(* Logix 5000 project; controller TFF vendor 1 type 14 code 107 rev 33.11; software revision 33.04; part 33 of 38 *)
(* tags used below, declared in another part *)
   Address : DINT;   // Temp Address
   Index : DINT;   // Index
   Index2 : DINT;   // Index
   result : DINT[2];
   SCL : SCALE;   // Scale Instruction
   AlarmAnalog : AlarmAnalog[50];   // Analog Alarm Array
   AlarmControl : AlarmControl;   // Alarm Control
   AnalogOutput : AnalogOutput[25];   // Analog Output Array
   AnalogPoint : AnalogInput[50];   // Analog Input Array
   DigitalInput : BOOL[256];   // Digital Input Array these bits are copied from Input cards.
   DigitalPoint : DigitalPoint[150];   // Digital Point Array
   ES001 : ALIAS FOR DigitalPoint[2];
   FlowPath : FlowPath[64];   // Flow Path Array
   FlowPathControl : FlowPathControl;   // Flow Path Control
   RawAnalogInputArray : INT[50];   // Array of analog input raw
   SysControl : SysControl;   // General system status and command
   Valve : Valve[100];   // Valve Array
   ValveControl : ValveControl;   // Valve Control
   ValveSwInput : BOOL[64];   // Valve digital input
(* Process, continued *)

ROUTINE modInputAnalog   (* ladder *)
// Analog Input Routine
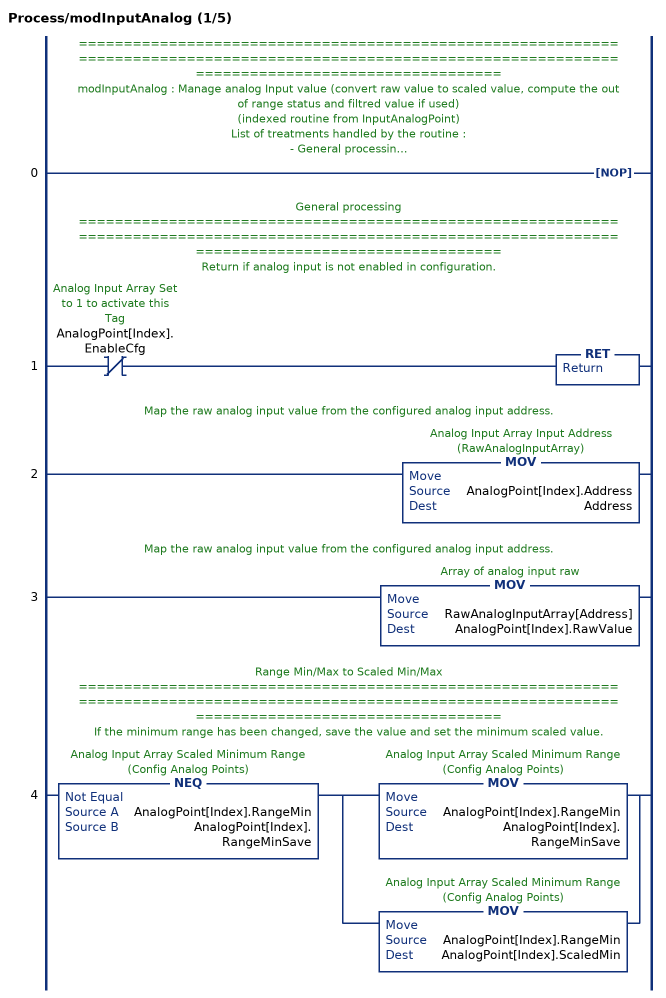
   // ==========================================================================================================================================================
   //                                            modInputAnalog : Manage analog Input value (convert raw value to scaled value, compute the out of range status and filtred value if used)
   //                                                                                                                        (indexed routine from InputAnalogPoint)
   //                                                     List of treatments handled by the routine :
   //                                                          - General processing
   //                                                          - Range Min/Max to Scaled Min/Max
   //                                                          - Out of Range status calculation
   //                                                          - filtering raw value
   //                                                          - Compute scaled value
   //                                                          - Map analog input value to alarm analog value
   //                                                     -----------------------------------------------------------------------------------------------------------------------------------------------------
   //                                                     History
   // 		2019-DEC-24 - Merck - Q. Spindler - Initial version for Candidate Release 1.00.00.00.a
   // 		2021-MAY-21 - Merck - Q. Spindler - Modifications for Candidate Release 1.00.00.00.e
   //                                                     - Out of Range status calculation, add exception for pressure sensors
   // ==========================================================================================================================================================
   0: NOP();
   // General processing
   // ==========================================================================================================================================================
   // Return if analog input is not enabled in configuration.
   1: XIO(AnalogPoint[Index].EnableCfg)RET();
   // Map the raw analog input value from the configured analog input address.
   2: MOV(AnalogPoint[Index].Address,Address);
   // Map the raw analog input value from the configured analog input address.
   3: MOV(RawAnalogInputArray[Address],AnalogPoint[Index].RawValue);
   // Range Min/Max to Scaled Min/Max
   // ==========================================================================================================================================================
   // If the minimum range has been changed, save the value and set the minimum scaled value.
   4: NEQ(AnalogPoint[Index].RangeMin,AnalogPoint[Index].RangeMinSave)[MOV(AnalogPoint[Index].RangeMin,AnalogPoint[Index].RangeMinSave) ,MOV(AnalogPoint[Index].RangeMin,AnalogPoint[Index].ScaledMin) ];
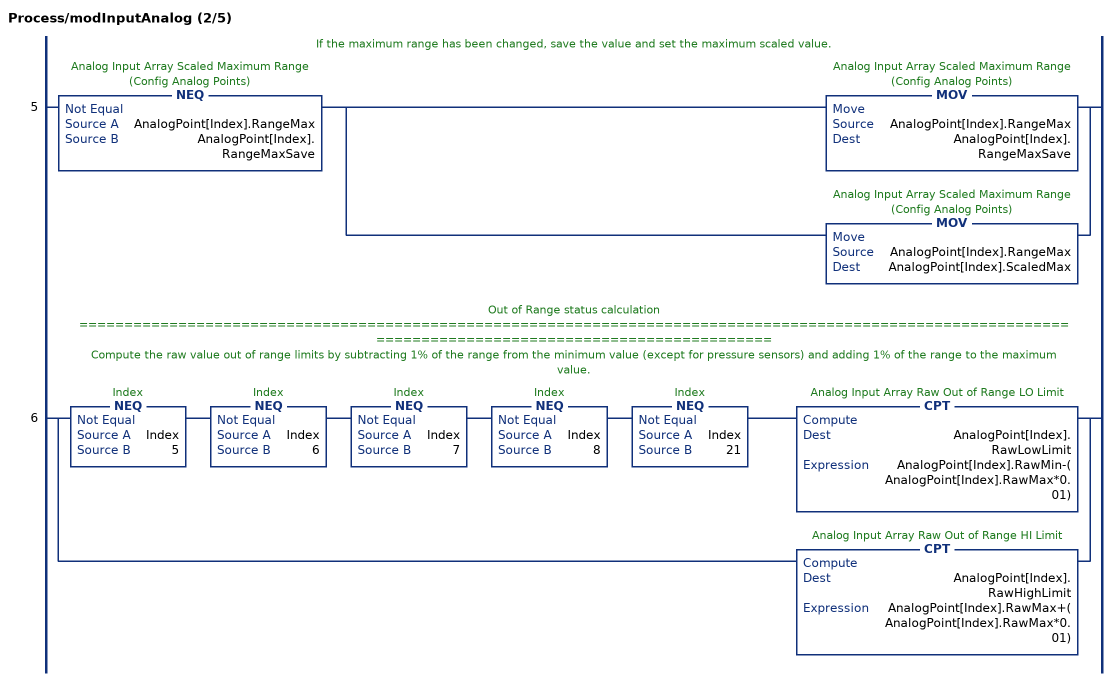
   // If the maximum range has been changed, save the value and set the maximum scaled value.
   5: NEQ(AnalogPoint[Index].RangeMax,AnalogPoint[Index].RangeMaxSave)[MOV(AnalogPoint[Index].RangeMax,AnalogPoint[Index].RangeMaxSave) ,MOV(AnalogPoint[Index].RangeMax,AnalogPoint[Index].ScaledMax) ];
   // Out of Range status calculation
   // ==========================================================================================================================================================
   // Compute the raw value out of range limits by subtracting 1% of the range from the minimum value (except for pressure sensors) and adding 1% of the range to the maximum value.
   6: [NEQ(Index,5) NEQ(Index,6) NEQ(Index,7) NEQ(Index,8) NEQ(Index,21) CPT(AnalogPoint[Index].RawLowLimit,AnalogPoint[Index].RawMin-(AnalogPoint[Index].RawMax*0.01)) ,CPT(AnalogPoint[Index].RawHighLimit,AnalogPoint[Index].RawMax+(AnalogPoint[Index].RawMax*0.01)) ];
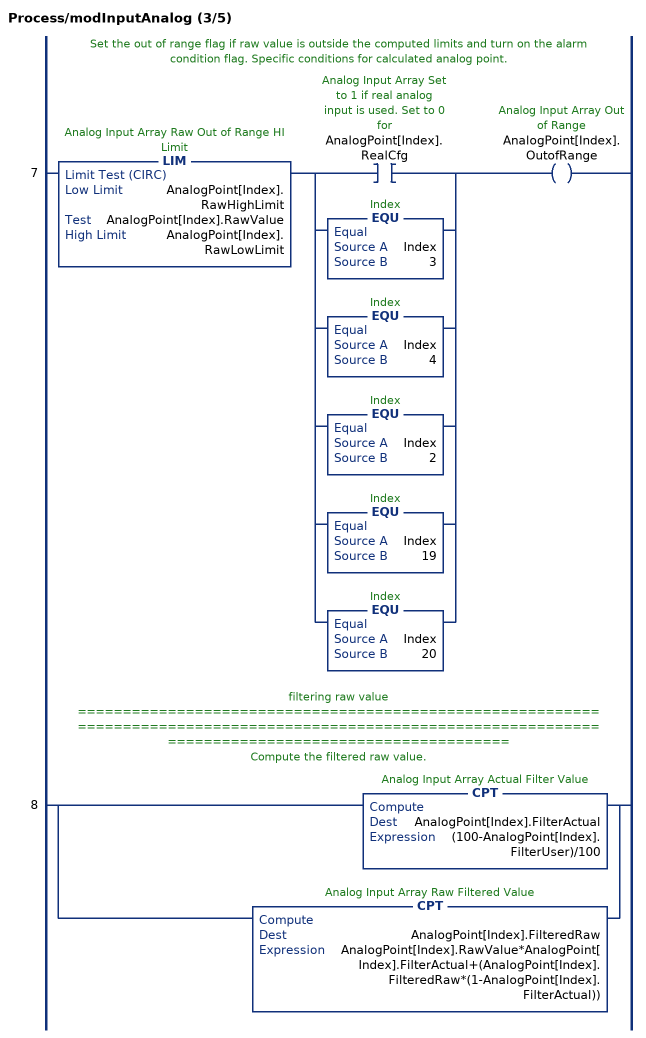
   // Set the out of range flag if raw value is outside the computed limits and turn on the alarm condition flag. Specific conditions for calculated analog point.
   7: LIM(AnalogPoint[Index].RawHighLimit,AnalogPoint[Index].RawValue,AnalogPoint[Index].RawLowLimit)[XIC(AnalogPoint[Index].RealCfg) ,EQU(Index,3) ,EQU(Index,4) ,EQU(Index,2) ,EQU(Index,19) ,EQU(Index,20) ]OTE(AnalogPoint[Index].OutofRange);
   // filtering raw value
   // ==========================================================================================================================================================
   // Compute the filtered raw value.
   8: [CPT(AnalogPoint[Index].FilterActual,(100-AnalogPoint[Index].FilterUser)/100) ,CPT(AnalogPoint[Index].FilteredRaw,AnalogPoint[Index].RawValue*AnalogPoint[Index].FilterActual+(AnalogPoint[Index].FilteredRaw*(1-AnalogPoint[Index].FilterActual))) ];
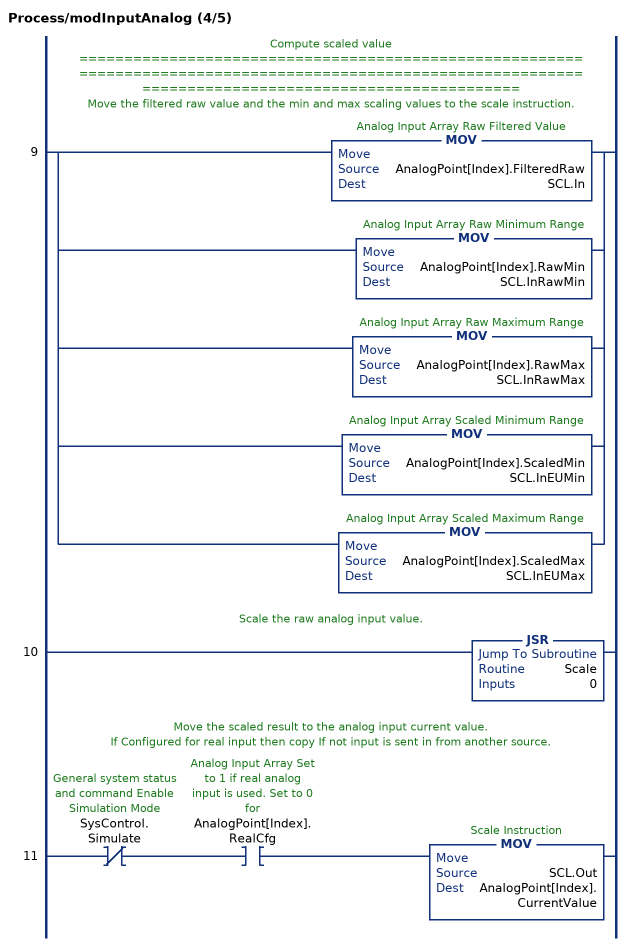
   // Compute scaled value
   // ==========================================================================================================================================================
   // Move the filtered raw value and the min and max scaling values to the scale instruction.
   9: [MOV(AnalogPoint[Index].FilteredRaw,SCL.In) ,MOV(AnalogPoint[Index].RawMin,SCL.InRawMin) ,MOV(AnalogPoint[Index].RawMax,SCL.InRawMax) ,MOV(AnalogPoint[Index].ScaledMin,SCL.InEUMin) ,MOV(AnalogPoint[Index].ScaledMax,SCL.InEUMax) ];
   // Scale the raw analog input value.
   10: JSR(Scale,0);
   // Move the scaled result to the analog input current value.
   // If Configured for real input then copy If not input is sent in from another source.
   11: XIO(SysControl.Simulate)XIC(AnalogPoint[Index].RealCfg)MOV(SCL.Out,AnalogPoint[Index].CurrentValue);
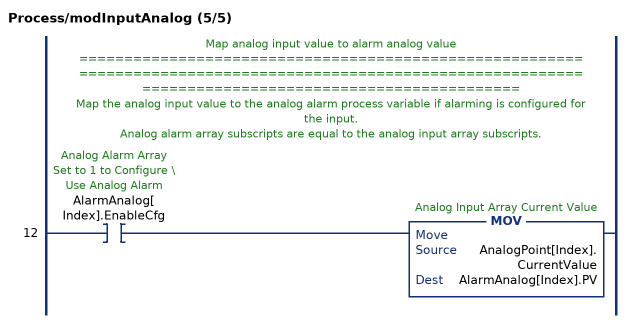
   // Map analog input value to alarm analog value
   // ==========================================================================================================================================================
   // Map the analog input value to the analog alarm process variable if alarming is configured for the input.
   // Analog alarm array subscripts are equal to the analog input array subscripts.
   12: XIC(AlarmAnalog[Index].EnableCfg)MOV(AnalogPoint[Index].CurrentValue,AlarmAnalog[Index].PV);
END_ROUTINE

ROUTINE modInputDigital   (* ladder *)
// Digital Input Routine
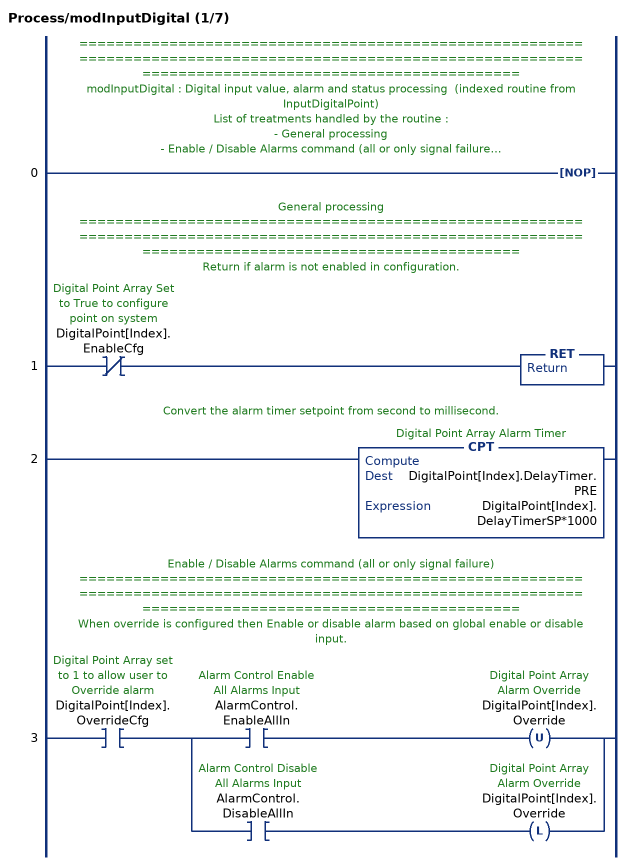
   // ==========================================================================================================================================================
   //                                                        modInputDigital : Digital input value, alarm and status processing  (indexed routine from InputDigitalPoint)
   //                                                     List of treatments handled by the routine :
   //                                                          - General processing
   //                                                          - Enable / Disable Alarms command (all or only signal failure)
   //                                                          - Digital alarm processing
   //                                                          - Digital input status
   //                                                          - Digital alarm status acknowledged
   //                                                          - Digital alarm status
   //                                                          - General processing
   //                                                          - Compute current value
   //                                                     -----------------------------------------------------------------------------------------------------------------------------------------------------
   //                                                     History
   // 		2019-DEC-24 - Merck - Q. Spindler - Initial version for Candidate Release 1.00.00.00.a
   // ==========================================================================================================================================================
   0: NOP();
   // General processing
   // ==========================================================================================================================================================
   // Return if alarm is not enabled in configuration.
   1: XIO(DigitalPoint[Index].EnableCfg)RET();
   // Convert the alarm timer setpoint from second to millisecond.
   2: CPT(DigitalPoint[Index].DelayTimer.PRE,DigitalPoint[Index].DelayTimerSP*1000);
   // Enable / Disable Alarms command (all or only signal failure)
   // ==========================================================================================================================================================
   // When override is configured then Enable or disable alarm based on global enable or disable input.
   3: XIC(DigitalPoint[Index].OverrideCfg)[XIC(AlarmControl.EnableAllIn) OTU(DigitalPoint[Index].Override) ,XIC(AlarmControl.DisableAllIn) OTL(DigitalPoint[Index].Override) ];
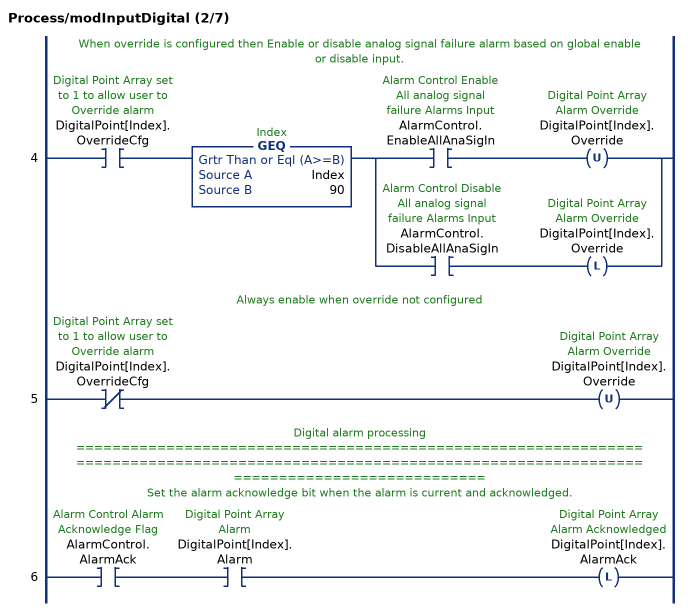
   // When override is configured then Enable or disable analog signal failure alarm based on global enable or disable input.
   4: XIC(DigitalPoint[Index].OverrideCfg)GEQ(Index,90)[XIC(AlarmControl.EnableAllAnaSigIn) OTU(DigitalPoint[Index].Override) ,XIC(AlarmControl.DisableAllAnaSigIn) OTL(DigitalPoint[Index].Override) ];
   // Always enable when override not configured
   5: XIO(DigitalPoint[Index].OverrideCfg)OTU(DigitalPoint[Index].Override);
   // Digital alarm processing
   // ==========================================================================================================================================================
   // Set the alarm acknowledge bit when the alarm is current and acknowledged.
   6: XIC(AlarmControl.AlarmAck)XIC(DigitalPoint[Index].Alarm)OTL(DigitalPoint[Index].AlarmAck);
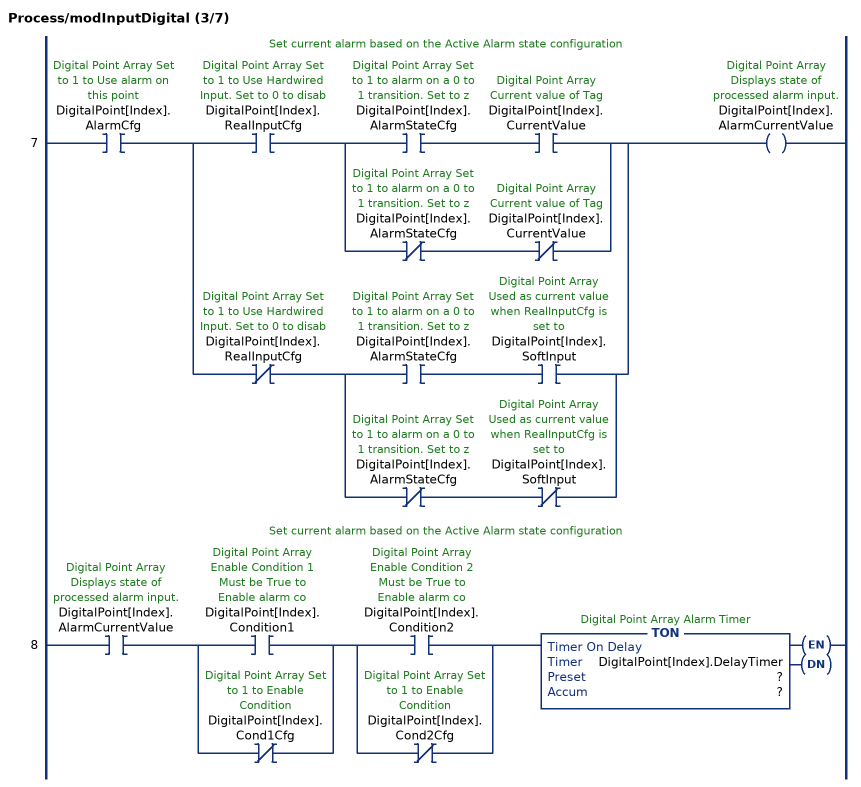
   // Set current alarm based on the Active Alarm state configuration
   7: XIC(DigitalPoint[Index].AlarmCfg)[XIC(DigitalPoint[Index].RealInputCfg) [XIC(DigitalPoint[Index].AlarmStateCfg) XIC(DigitalPoint[Index].CurrentValue) ,XIO(DigitalPoint[Index].AlarmStateCfg) XIO(DigitalPoint[Index].CurrentValue) ] ,XIO(DigitalPoint[Index].RealInputCfg) [XIC(DigitalPoint[Index].AlarmStateCfg) XIC(DigitalPoint[Index].SoftInput) ,XIO(DigitalPoint[Index].AlarmStateCfg) XIO(DigitalPoint[Index].SoftInput) ] ]OTE(DigitalPoint[Index].AlarmCurrentValue);
   // Set current alarm based on the Active Alarm state configuration
   8: XIC(DigitalPoint[Index].AlarmCurrentValue)[XIC(DigitalPoint[Index].Condition1) ,XIO(DigitalPoint[Index].Cond1Cfg) ][XIC(DigitalPoint[Index].Condition2) ,XIO(DigitalPoint[Index].Cond2Cfg) ]TON(DigitalPoint[Index].DelayTimer,?,?);
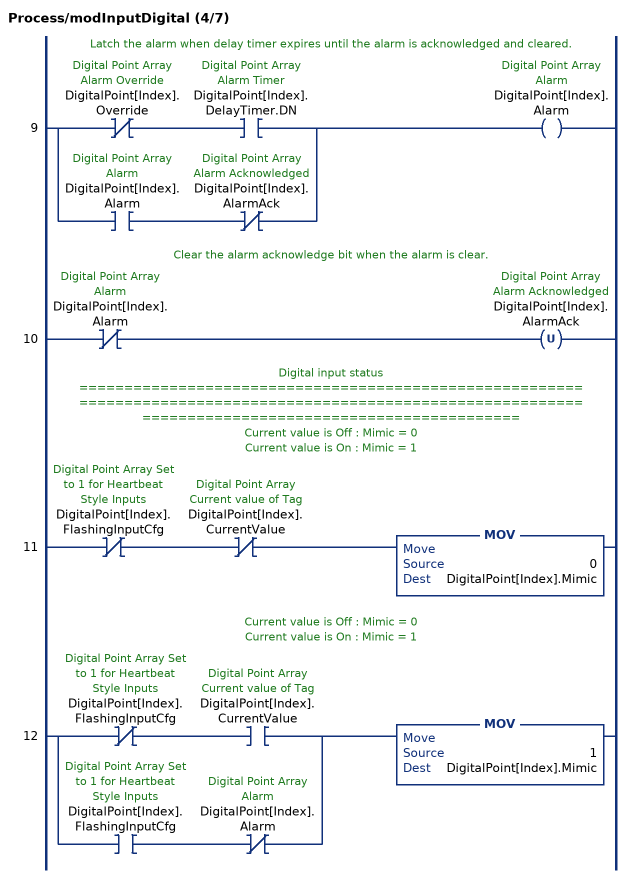
   // Latch the alarm when delay timer expires until the alarm is acknowledged and cleared.
   9: [XIO(DigitalPoint[Index].Override) XIC(DigitalPoint[Index].DelayTimer.DN) ,XIC(DigitalPoint[Index].Alarm) XIO(DigitalPoint[Index].AlarmAck) ]OTE(DigitalPoint[Index].Alarm);
   // Clear the alarm acknowledge bit when the alarm is clear.
   10: XIO(DigitalPoint[Index].Alarm)OTU(DigitalPoint[Index].AlarmAck);
   // Digital input status
   // ==========================================================================================================================================================
   // Current value is Off : Mimic = 0
   // Current value is On : Mimic = 1
   11: XIO(DigitalPoint[Index].FlashingInputCfg)XIO(DigitalPoint[Index].CurrentValue)MOV(0,DigitalPoint[Index].Mimic);
   // Current value is Off : Mimic = 0
   // Current value is On : Mimic = 1
   12: [XIO(DigitalPoint[Index].FlashingInputCfg) XIC(DigitalPoint[Index].CurrentValue) ,XIC(DigitalPoint[Index].FlashingInputCfg) XIO(DigitalPoint[Index].Alarm) ]MOV(1,DigitalPoint[Index].Mimic);
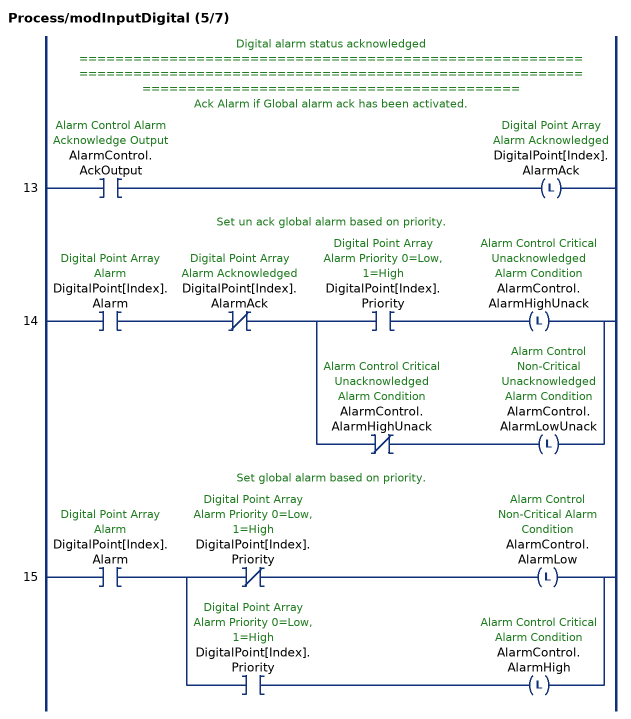
   // Digital alarm status acknowledged
   // ==========================================================================================================================================================
   // Ack Alarm if Global alarm ack has been activated.
   13: XIC(AlarmControl.AckOutput)OTL(DigitalPoint[Index].AlarmAck);
   // Set un ack global alarm based on priority.
   14: XIC(DigitalPoint[Index].Alarm)XIO(DigitalPoint[Index].AlarmAck)[XIC(DigitalPoint[Index].Priority) OTL(AlarmControl.AlarmHighUnack) ,XIO(AlarmControl.AlarmHighUnack) OTL(AlarmControl.AlarmLowUnack) ];
   // Set global alarm based on priority.
   15: XIC(DigitalPoint[Index].Alarm)[XIO(DigitalPoint[Index].Priority) OTL(AlarmControl.AlarmLow) ,XIC(DigitalPoint[Index].Priority) OTL(AlarmControl.AlarmHigh) ];
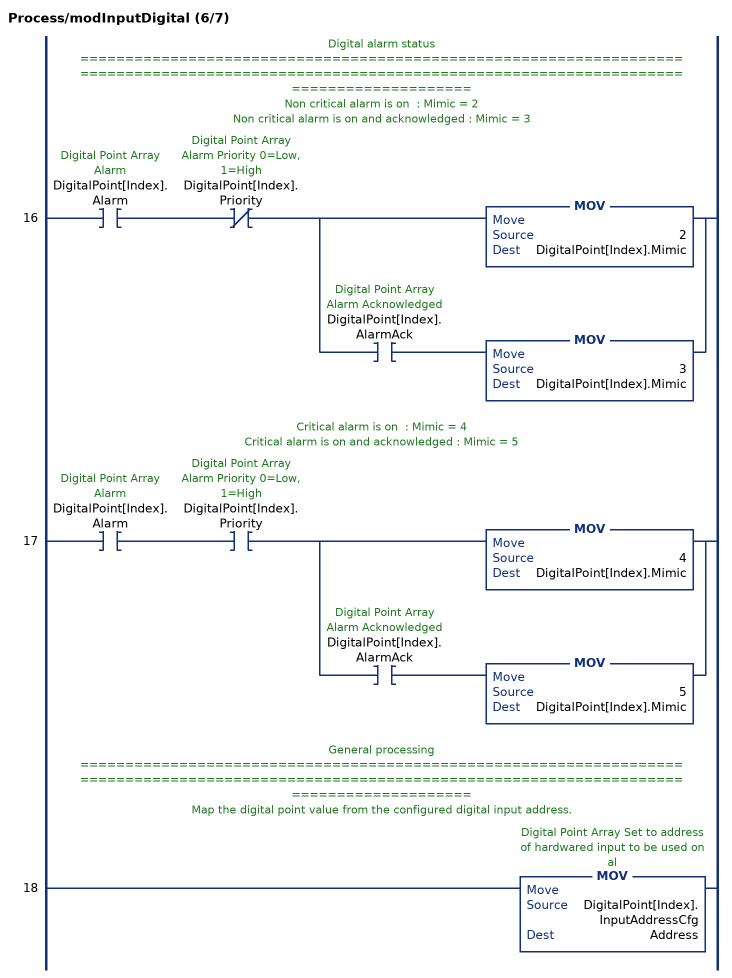
   // Digital alarm status
   // ==========================================================================================================================================================
   // Non critical alarm is on  : Mimic = 2
   // Non critical alarm is on and acknowledged : Mimic = 3
   16: XIC(DigitalPoint[Index].Alarm)XIO(DigitalPoint[Index].Priority)[MOV(2,DigitalPoint[Index].Mimic) ,XIC(DigitalPoint[Index].AlarmAck) MOV(3,DigitalPoint[Index].Mimic) ];
   // Critical alarm is on  : Mimic = 4
   // Critical alarm is on and acknowledged : Mimic = 5
   17: XIC(DigitalPoint[Index].Alarm)XIC(DigitalPoint[Index].Priority)[MOV(4,DigitalPoint[Index].Mimic) ,XIC(DigitalPoint[Index].AlarmAck) MOV(5,DigitalPoint[Index].Mimic) ];
   // General processing
   // ==========================================================================================================================================================
   // Map the digital point value from the configured digital input address.
   18: MOV(DigitalPoint[Index].InputAddressCfg,Address);
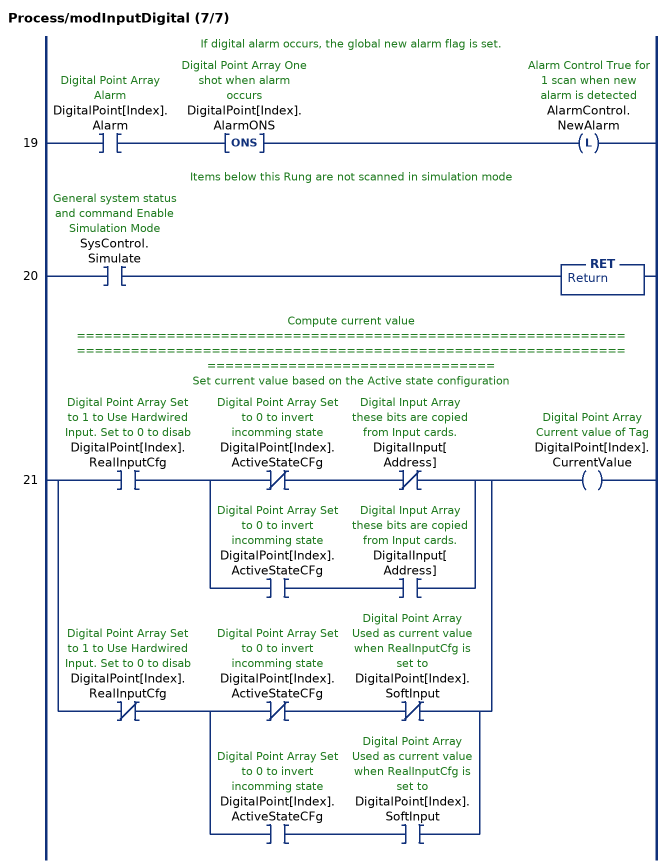
   // If digital alarm occurs, the global new alarm flag is set.
   19: XIC(DigitalPoint[Index].Alarm)ONS(DigitalPoint[Index].AlarmONS)OTL(AlarmControl.NewAlarm);
   // Items below this Rung are not scanned in simulation mode
   20: XIC(SysControl.Simulate)RET();
   // Compute current value
   // ==========================================================================================================================================================
   // Set current value based on the Active state configuration
   21: [XIC(DigitalPoint[Index].RealInputCfg) [XIO(DigitalPoint[Index].ActiveStateCFg) XIO(DigitalInput[Address]) ,XIC(DigitalPoint[Index].ActiveStateCFg) XIC(DigitalInput[Address]) ] ,XIO(DigitalPoint[Index].RealInputCfg) [XIO(DigitalPoint[Index].ActiveStateCFg) XIO(DigitalPoint[Index].SoftInput) ,XIC(DigitalPoint[Index].ActiveStateCFg) XIC(DigitalPoint[Index].SoftInput) ] ]OTE(DigitalPoint[Index].CurrentValue);
END_ROUTINE

ROUTINE modOutputAnalog   (* ladder *)
// Analog Output Routine
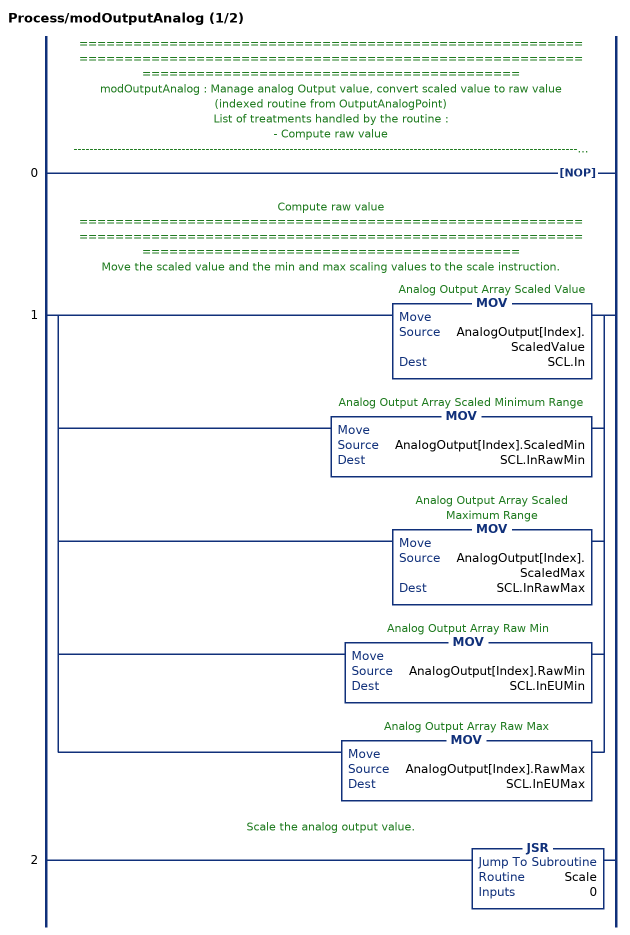
   // ==========================================================================================================================================================
   //                                            modOutputAnalog : Manage analog Output value, convert scaled value to raw value (indexed routine from OutputAnalogPoint)
   //                                                     List of treatments handled by the routine :
   //                                                          - Compute raw value
   //                                                     -----------------------------------------------------------------------------------------------------------------------------------------------------
   //                                                     History
   // 		2019-DEC-24 - Merck - Q. Spindler - Initial version for Candidate Release 1.00.00.00.a
   // ==========================================================================================================================================================
   0: NOP();
   // Compute raw value
   // ==========================================================================================================================================================
   // Move the scaled value and the min and max scaling values to the scale instruction.
   1: [MOV(AnalogOutput[Index].ScaledValue,SCL.In) ,MOV(AnalogOutput[Index].ScaledMin,SCL.InRawMin) ,MOV(AnalogOutput[Index].ScaledMax,SCL.InRawMax) ,MOV(AnalogOutput[Index].RawMin,SCL.InEUMin) ,MOV(AnalogOutput[Index].RawMax,SCL.InEUMax) ];
   // Scale the analog output value.
   2: JSR(Scale,0);
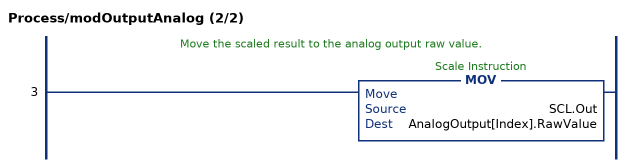
   // Move the scaled result to the analog output raw value.
   3: MOV(SCL.Out,AnalogOutput[Index].RawValue);
END_ROUTINE

ROUTINE ModValveControl   (* ladder *)
// Valve Control Routine
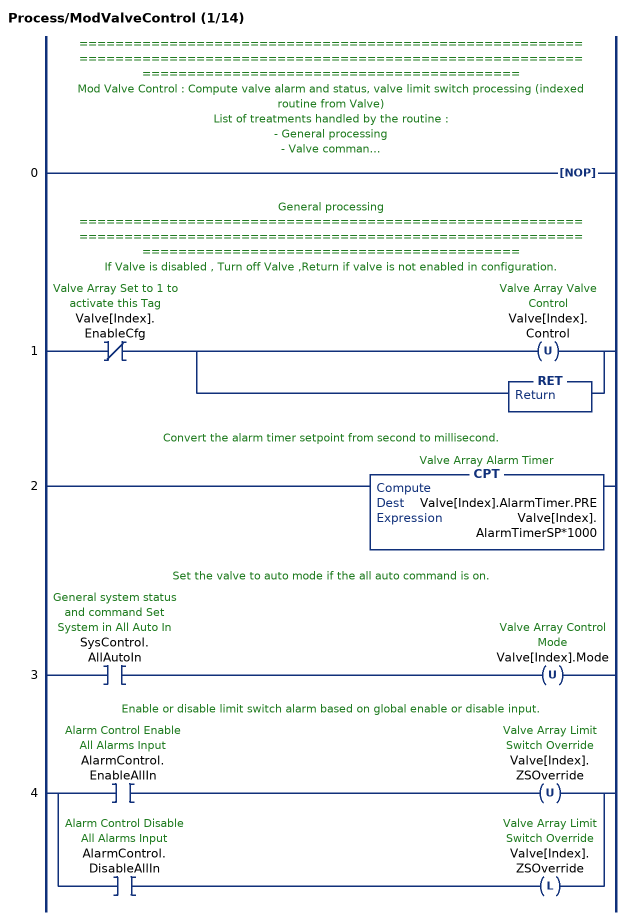
   // ==========================================================================================================================================================
   //                                                      Mod Valve Control : Compute valve alarm and status, valve limit switch processing (indexed routine from Valve)
   //                                                     List of treatments handled by the routine :
   //                                                          - General processing
   //                                                          - Valve command
   //                                                          - Valve limit switch
   //                                                          - Valve status
   //                                                          - Valve alarm
   //                                                          - Valve alarm status
   //                                                          - Valve status for flowpath logic
   //                                                          - Output command
   //                                                     -----------------------------------------------------------------------------------------------------------------------------------------------------
   //                                                     History
   // 		2019-DEC-24 - Merck - Q. Spindler - Initial version for Candidate Release 1.00.00.00.a
   // ==========================================================================================================================================================
   0: NOP();
   // General processing
   // ==========================================================================================================================================================
   // If Valve is disabled , Turn off Valve ,Return if valve is not enabled in configuration.
   1: XIO(Valve[Index].EnableCfg)[OTU(Valve[Index].Control) ,RET() ];
   // Convert the alarm timer setpoint from second to millisecond.
   2: CPT(Valve[Index].AlarmTimer.PRE,Valve[Index].AlarmTimerSP*1000);
   // Set the valve to auto mode if the all auto command is on.
   3: XIC(SysControl.AllAutoIn)OTU(Valve[Index].Mode);
   // Enable or disable limit switch alarm based on global enable or disable input.
   4: [XIC(AlarmControl.EnableAllIn) OTU(Valve[Index].ZSOverride) ,XIC(AlarmControl.DisableAllIn) OTL(Valve[Index].ZSOverride) ];
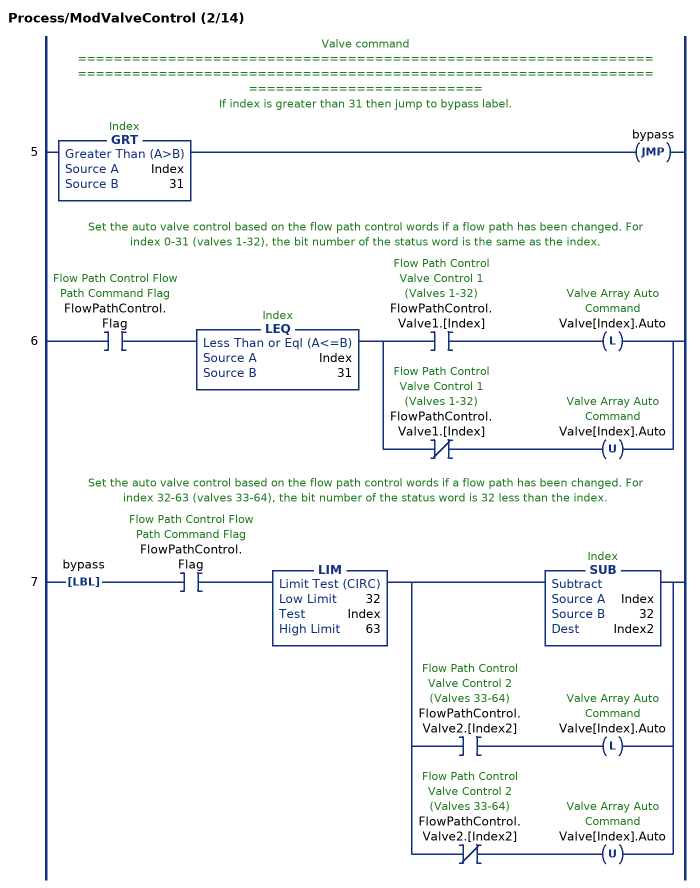
   // Valve command
   // ==========================================================================================================================================================
   // If index is greater than 31 then jump to bypass label.
   5: GRT(Index,31)JMP(bypass);
   // Set the auto valve control based on the flow path control words if a flow path has been changed. For index 0-31 (valves 1-32), the bit number of the status word is the same as the index.
   6: XIC(FlowPathControl.Flag)LEQ(Index,31)[XIC(FlowPathControl.Valve1.[Index]) OTL(Valve[Index].Auto) ,XIO(FlowPathControl.Valve1.[Index]) OTU(Valve[Index].Auto) ];
   // Set the auto valve control based on the flow path control words if a flow path has been changed. For index 32-63 (valves 33-64), the bit number of the status word is 32 less than the index.
   7: LBL(bypass)XIC(FlowPathControl.Flag)LIM(32,Index,63)[SUB(Index,32,Index2) ,XIC(FlowPathControl.Valve2.[Index2]) OTL(Valve[Index].Auto) ,XIO(FlowPathControl.Valve2.[Index2]) OTU(Valve[Index].Auto) ];
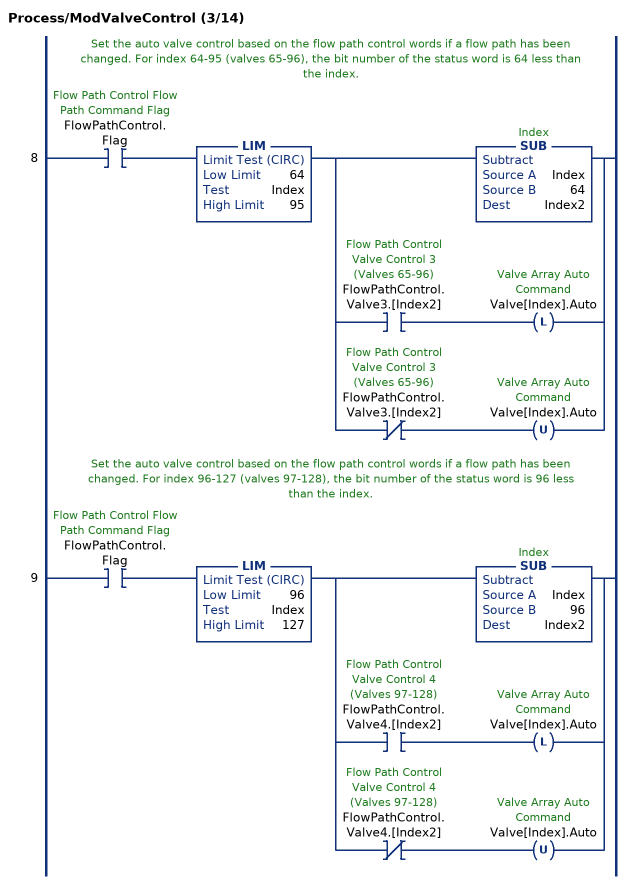
   // Set the auto valve control based on the flow path control words if a flow path has been changed. For index 64-95 (valves 65-96), the bit number of the status word is 64 less than the index.
   8: XIC(FlowPathControl.Flag)LIM(64,Index,95)[SUB(Index,64,Index2) ,XIC(FlowPathControl.Valve3.[Index2]) OTL(Valve[Index].Auto) ,XIO(FlowPathControl.Valve3.[Index2]) OTU(Valve[Index].Auto) ];
   // Set the auto valve control based on the flow path control words if a flow path has been changed. For index 96-127 (valves 97-128), the bit number of the status word is 96 less than the index.
   9: XIC(FlowPathControl.Flag)LIM(96,Index,127)[SUB(Index,96,Index2) ,XIC(FlowPathControl.Valve4.[Index2]) OTL(Valve[Index].Auto) ,XIO(FlowPathControl.Valve4.[Index2]) OTU(Valve[Index].Auto) ];
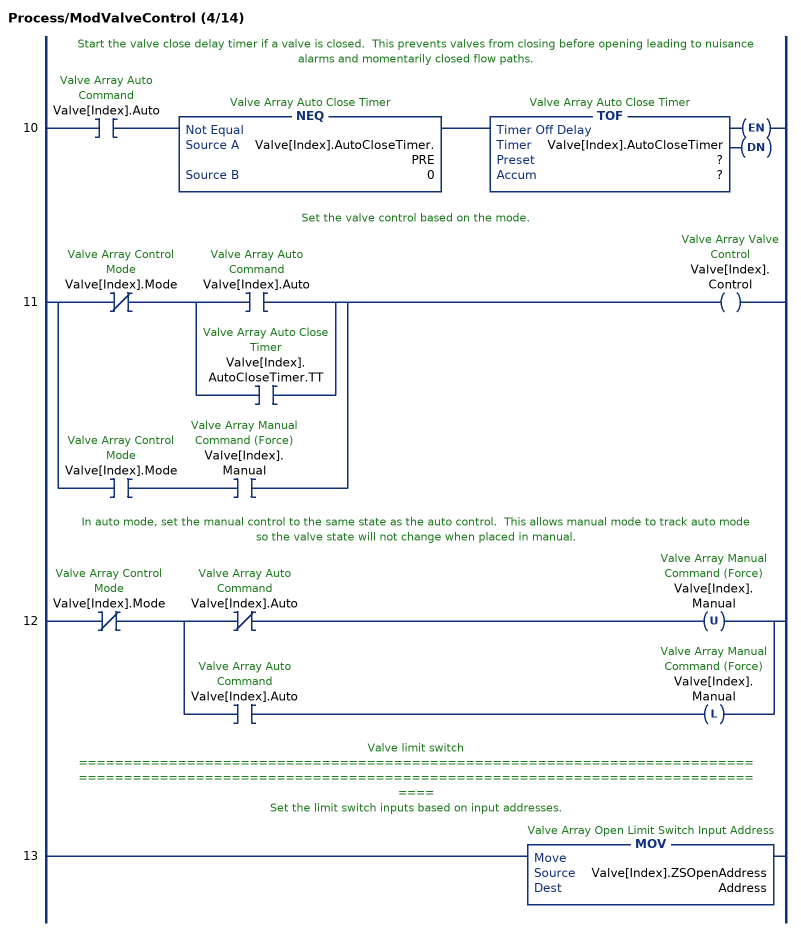
   // Start the valve close delay timer if a valve is closed.  This prevents valves from closing before opening leading to nuisance alarms and momentarily closed flow paths.
   10: XIC(Valve[Index].Auto)NEQ(Valve[Index].AutoCloseTimer.PRE,0)TOF(Valve[Index].AutoCloseTimer,?,?);
   // Set the valve control based on the mode.
   11: [XIO(Valve[Index].Mode) [XIC(Valve[Index].Auto) ,XIC(Valve[Index].AutoCloseTimer.TT) ] ,XIC(Valve[Index].Mode) XIC(Valve[Index].Manual) ]OTE(Valve[Index].Control);
   // In auto mode, set the manual control to the same state as the auto control.  This allows manual mode to track auto mode so the valve state will not change when placed in manual.
   12: XIO(Valve[Index].Mode)[XIO(Valve[Index].Auto) OTU(Valve[Index].Manual) ,XIC(Valve[Index].Auto) OTL(Valve[Index].Manual) ];
   // Valve limit switch
   // ==========================================================================================================================================================
   // Set the limit switch inputs based on input addresses.
   13: MOV(Valve[Index].ZSOpenAddress,Address);
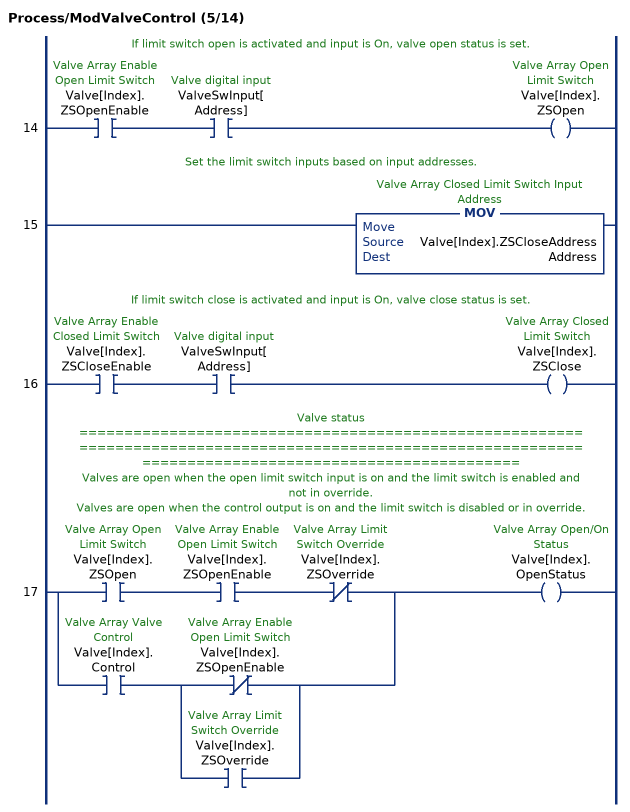
   // If limit switch open is activated and input is On, valve open status is set.
   14: XIC(Valve[Index].ZSOpenEnable)XIC(ValveSwInput[Address])OTE(Valve[Index].ZSOpen);
   // Set the limit switch inputs based on input addresses.
   15: MOV(Valve[Index].ZSCloseAddress,Address);
   // If limit switch close is activated and input is On, valve close status is set.
   16: XIC(Valve[Index].ZSCloseEnable)XIC(ValveSwInput[Address])OTE(Valve[Index].ZSClose);
   // Valve status
   // ==========================================================================================================================================================
   // Valves are open when the open limit switch input is on and the limit switch is enabled and not in override.
   // Valves are open when the control output is on and the limit switch is disabled or in override.
   17: [XIC(Valve[Index].ZSOpen) XIC(Valve[Index].ZSOpenEnable) XIO(Valve[Index].ZSOverride) ,XIC(Valve[Index].Control) [XIO(Valve[Index].ZSOpenEnable) ,XIC(Valve[Index].ZSOverride) ] ]OTE(Valve[Index].OpenStatus);
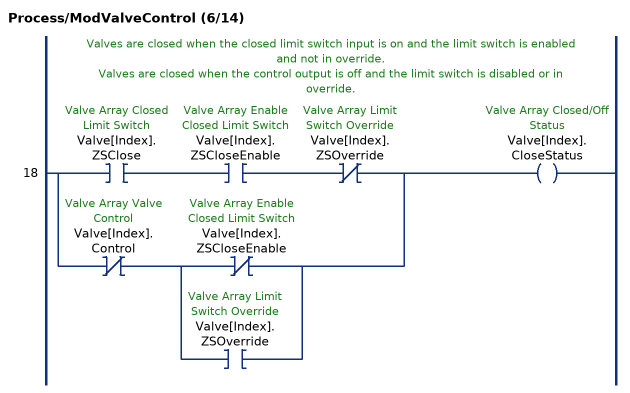
   // Valves are closed when the closed limit switch input is on and the limit switch is enabled and not in override.
   // Valves are closed when the control output is off and the limit switch is disabled or in override.
   18: [XIC(Valve[Index].ZSClose) XIC(Valve[Index].ZSCloseEnable) XIO(Valve[Index].ZSOverride) ,XIO(Valve[Index].Control) [XIO(Valve[Index].ZSCloseEnable) ,XIC(Valve[Index].ZSOverride) ] ]OTE(Valve[Index].CloseStatus);
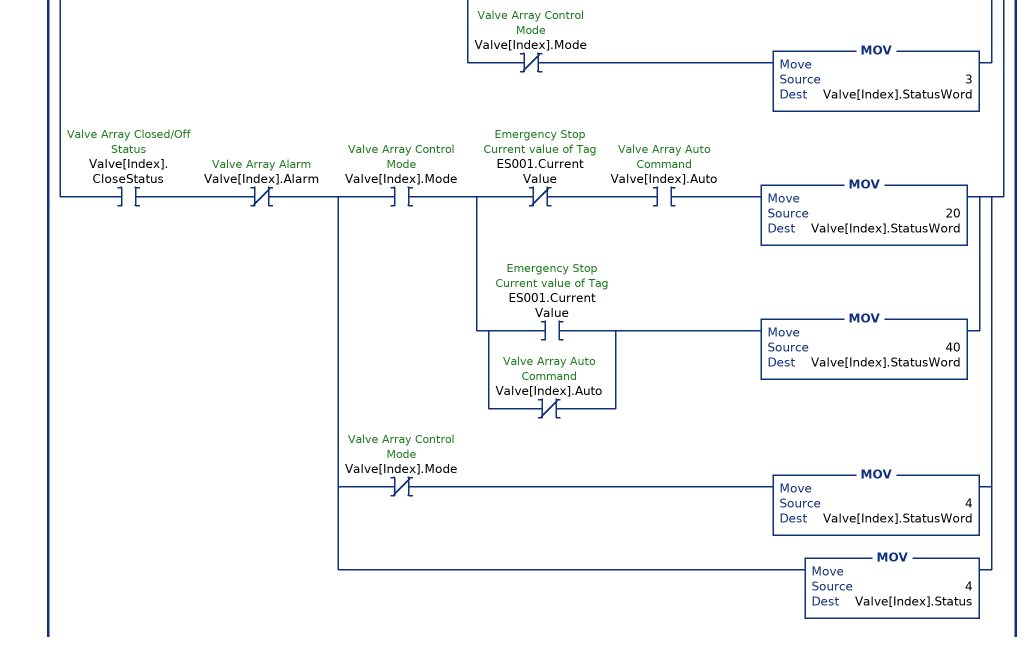
   // Auto Valve Status Word.
   // 1 = Travel (Auto Mode) , 10 = Travel (Manual Mode)
   // 2 = Open/On (Auto Mode) , 20 = Open/On (Manual Mode)
   // 3 = Travel (Auto Mode) , 30 = Travel (Manual Mode)
   // 4 = Closed/Off (Auto Mode) , 40 = Closed/Off (Manual Mode)
   // If the option VlvPstnSensor is disabled, Open/On and Closed/Off are inverted if an Emergency Stop is triggered to correspond to the physical state (state without pressure)
   19: [XIO(Valve[Index].OpenStatus) XIO(Valve[Index].CloseStatus) XIO(Valve[Index].Alarm) [XIC(Valve[Index].Mode) MOV(10,Valve[Index].StatusWord) ,XIO(Valve[Index].Mode) MOV(1,Valve[Index].StatusWord) ] ,XIC(Valve[Index].OpenStatus) XIO(Valve[Index].Alarm) [XIC(Valve[Index].Mode) [XIO(ES001.CurrentValue) XIO(Valve[Index].Auto) MOV(40,Valve[Index].StatusWord) ,[XIC(ES001.CurrentValue) ,XIC(Valve[Index].Auto) ] MOV(20,Valve[Index].StatusWord) ] ,XIO(Valve[Index].Mode) MOV(2,Valve[Index].StatusWord) ,MOV(2,Valve[Index].Status) ] ,XIC(Valve[Index].OpenStatus) XIC(Valve[Index].CloseStatus) XIO(Valve[Index].Alarm) [XIC(Valve[Index].Mode) MOV(30,Valve[Index].StatusWord) ,XIO(Valve[Index].Mode) MOV(3,Valve[Index].StatusWord) ] ,XIC(Valve[Index].CloseStatus) XIO(Valve[Index].Alarm) [XIC(Valve[Index].Mode) [XIO(ES001.CurrentValue) XIC(Valve[Index].Auto) MOV(20,Valve[Index].StatusWord) ,[XIC(ES001.CurrentValue) ,XIO(Valve[Index].Auto) ] MOV(40,Valve[Index].StatusWord) ] ,XIO(Valve[Index].Mode) MOV(4,Valve[Index].StatusWord) ,MOV(4,Valve[Index].Status) ] ];
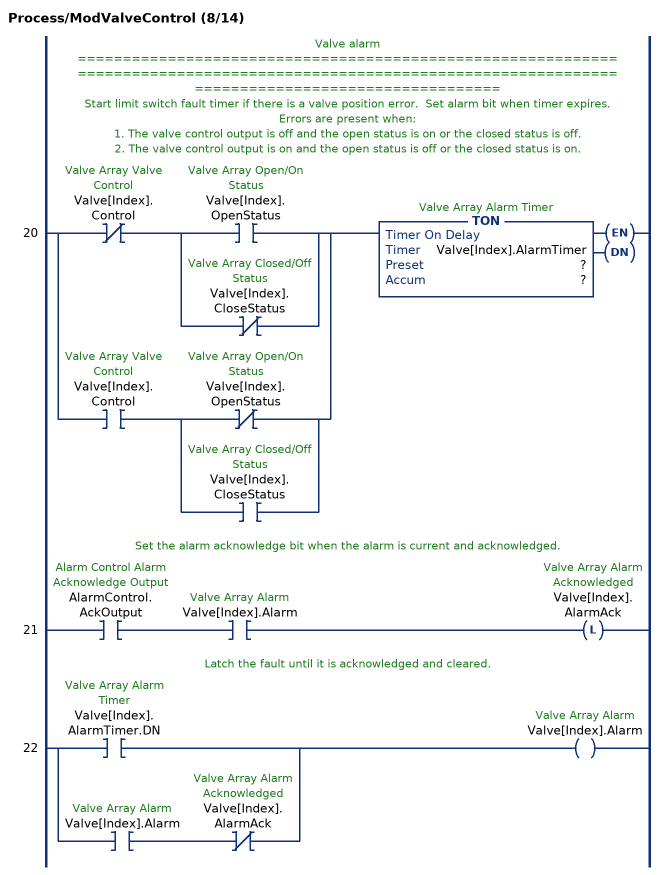
   // Valve alarm
   // ==========================================================================================================================================================
   // Start limit switch fault timer if there is a valve position error.  Set alarm bit when timer expires.
   // Errors are present when:
   // 1. The valve control output is off and the open status is on or the closed status is off.
   // 2. The valve control output is on and the open status is off or the closed status is on.
   20: [XIO(Valve[Index].Control) [XIC(Valve[Index].OpenStatus) ,XIO(Valve[Index].CloseStatus) ] ,XIC(Valve[Index].Control) [XIO(Valve[Index].OpenStatus) ,XIC(Valve[Index].CloseStatus) ] ]TON(Valve[Index].AlarmTimer,?,?);
   // Set the alarm acknowledge bit when the alarm is current and acknowledged.
   21: XIC(AlarmControl.AckOutput)XIC(Valve[Index].Alarm)OTL(Valve[Index].AlarmAck);
   // Latch the fault until it is acknowledged and cleared.
   22: [XIC(Valve[Index].AlarmTimer.DN) ,XIC(Valve[Index].Alarm) XIO(Valve[Index].AlarmAck) ]OTE(Valve[Index].Alarm);
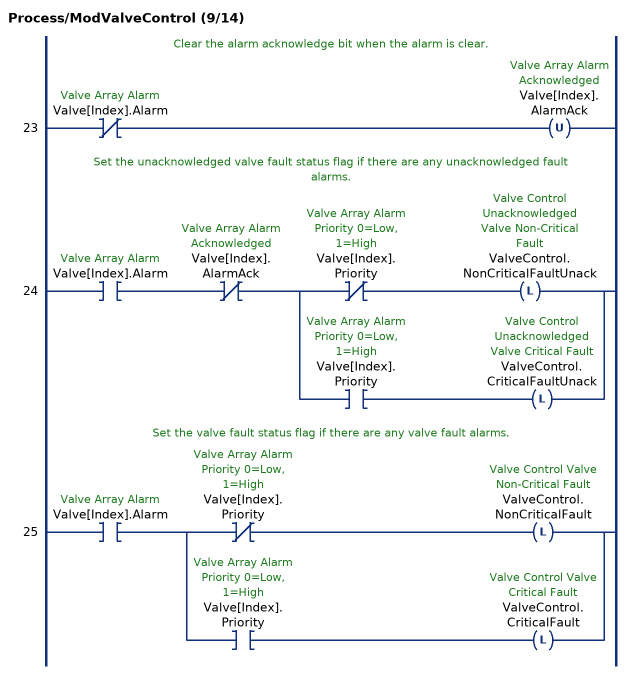
   // Clear the alarm acknowledge bit when the alarm is clear.
   23: XIO(Valve[Index].Alarm)OTU(Valve[Index].AlarmAck);
   // Set the unacknowledged valve fault status flag if there are any unacknowledged fault alarms.
   24: XIC(Valve[Index].Alarm)XIO(Valve[Index].AlarmAck)[XIO(Valve[Index].Priority) OTL(ValveControl.NonCriticalFaultUnack) ,XIC(Valve[Index].Priority) OTL(ValveControl.CriticalFaultUnack) ];
   // Set the valve fault status flag if there are any valve fault alarms.
   25: XIC(Valve[Index].Alarm)[XIO(Valve[Index].Priority) OTL(ValveControl.NonCriticalFault) ,XIC(Valve[Index].Priority) OTL(ValveControl.CriticalFault) ];
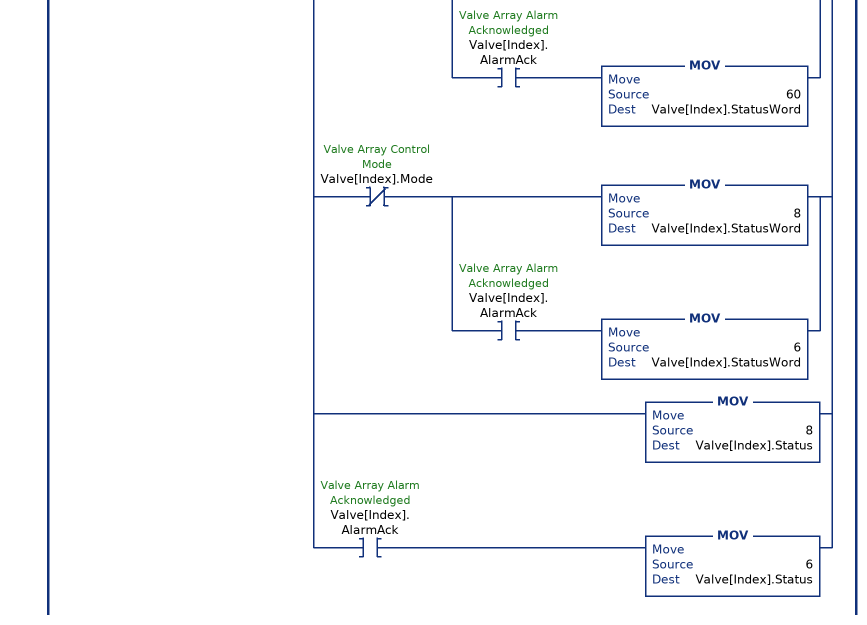
   // Valve alarm status
   // ==========================================================================================================================================================
   // Auto Valve Status Word, based on priority if any Vavle alarms..
   // 5 = Non Critical Alarm (Auto Mode) , 50 = Non Critical Alarm (Manual Mode)
   // 6 = Critical Alarm (Auto Mode) , 60 = Critical Alarm (Manual Mode)
   // 7 = Non Critical Alarm Unack (Auto Mode) , 70 = Non Critical Alarm Unack  (Manual Mode)
   // 8 = Critical Alarm Unack (Auto Mode) , 80 = Critical Alarm Unack  (Manual Mode)
   26: XIC(Valve[Index].Alarm)[XIO(Valve[Index].Priority) [XIC(Valve[Index].Mode) [MOV(70,Valve[Index].StatusWord) ,XIC(Valve[Index].AlarmAck) MOV(50,Valve[Index].StatusWord) ] ,XIO(Valve[Index].Mode) [MOV(7,Valve[Index].StatusWord) ,XIC(Valve[Index].AlarmAck) MOV(5,Valve[Index].StatusWord) ] ,[MOV(7,Valve[Index].Status) ,XIC(Valve[Index].AlarmAck) MOV(5,Valve[Index].Status) ] ] ,XIC(Valve[Index].Priority) [XIC(Valve[Index].Mode) [MOV(80,Valve[Index].StatusWord) ,XIC(Valve[Index].AlarmAck) MOV(60,Valve[Index].StatusWord) ] ,XIO(Valve[Index].Mode) [MOV(8,Valve[Index].StatusWord) ,XIC(Valve[Index].AlarmAck) MOV(6,Valve[Index].StatusWord) ] ,[MOV(8,Valve[Index].Status) ,XIC(Valve[Index].AlarmAck) MOV(6,Valve[Index].Status) ] ] ];
